Staubli VAL3: HMI_message.dtx

bool bToHome
string sRobotMsg[40]
bool bBack
num nMsgType
string sCurrentMsg
